(* IEC 61131-3 sources: llm-plc-st-eval/data/processed_definitivo/gemini-3.1-pro-preview/I8/zero_shot, 3 files *)

(* ---- ejec_1.st ---- *)
FUNCTION_BLOCK FB_Compresor
VAR_INPUT
    pOilOk    : BOOL; // Presión de aceite correcta
    tempOk    : BOOL; // Temperatura correcta
    sinAlm    : BOOL; // Ausencia de alarmas
    btnMarcha : BOOL; // Botón de arranque
    btnParo   : BOOL; // Botón de detención
END_VAR

VAR_OUTPUT
    comp         : BOOL; // Comando de marcha del compresor
    causaBloqueo : INT;  // Código del permisivo faltante (0=Ninguno, 1=Aceite, 2=Temp, 3=Alarma)
END_VAR

VAR
    timerOil   : TON;    // Temporizador para validar la presión de aceite
    edgeMarcha : R_TRIG; // Detector de flanco de subida para el botón de marcha
    permisivos : BOOL;   // Bandera interna de todos los permisivos OK
END_VAR

// 1. Evaluación del tiempo de la presión de aceite (3 segundos continuos)
timerOil(IN := pOilOk, PT := T#3S);

// 2. Determinación de la causa de bloqueo (Prioridad al número menor)
IF NOT timerOil.Q THEN
    causaBloqueo := 1; // Falta presión de aceite o no ha transcurrido el tiempo
ELSIF NOT tempOk THEN
    causaBloqueo := 2; // Falta temperatura correcta
ELSIF NOT sinAlm THEN
    causaBloqueo := 3; // Presencia de alarma
ELSE
    causaBloqueo := 0; // Todos los permisivos se cumplen
END_IF;

// 3. Consolidación de permisivos
permisivos := (causaBloqueo = 0);

// 4. Detección de la pulsación de marcha (transición FALSE a TRUE)
edgeMarcha(CLK := btnMarcha);

// 5. Lógica de arranque y paro del compresor
// El paro y la pérdida de permisivos tienen prioridad absoluta
IF btnParo OR NOT permisivos THEN
    comp := FALSE;
// Solo arranca con un nuevo flanco de subida si los permisivos están listos
ELSIF edgeMarcha.Q AND permisivos THEN
    comp := TRUE;
END_IF;

END_FUNCTION_BLOCK

(* ---- ejec_2.st ---- *)
FUNCTION_BLOCK FB_Compresor
VAR_INPUT
    pOilOk    : BOOL; // Presión de aceite correcta
    tempOk    : BOOL; // Temperatura correcta
    sinAlm    : BOOL; // Ausencia de alarmas
    btnMarcha : BOOL; // Botón de arranque
    btnParo   : BOOL; // Botón de parada
END_VAR

VAR_OUTPUT
    comp         : BOOL; // Comando de arranque del compresor
    causaBloqueo : INT;  // Código del permisivo faltante (0=Ninguno, 1=Aceite, 2=Temp, 3=Alarma)
END_VAR

VAR
    tonOil     : TON;    // Temporizador para validar la presión de aceite
    trigMarcha : R_TRIG; // Detector de flanco de subida para el arranque
    permisivos : BOOL;   // Marca interna de todos los permisivos cumplidos
END_VAR

// 1. Temporizador: requiere 3 segundos continuos de pOilOk
tonOil(IN := pOilOk, PT := T#3S);

// 2. Lógica de diagnóstico de bloqueo (prioridad al número menor mediante IF-ELSIF)
IF NOT tonOil.Q THEN
    causaBloqueo := 1; // Falla 1: Presión de aceite no establecida
ELSIF NOT tempOk THEN
    causaBloqueo := 2; // Falla 2: Temperatura incorrecta
ELSIF NOT sinAlm THEN
    causaBloqueo := 3; // Falla 3: Alarma activa
ELSE
    causaBloqueo := 0; // Sin fallas: Todos los permisivos OK
END_IF;

// 3. Evaluación global de permisivos
permisivos := (causaBloqueo = 0);

// 4. Detección de pulsación (transición FALSE a TRUE) del botón de marcha
trigMarcha(CLK := btnMarcha);

// 5. Lógica de control de marcha/paro del compresor
IF btnParo OR NOT permisivos THEN
    // El paro y la pérdida de permisivos tienen prioridad y detienen el equipo
    comp := FALSE;
ELSIF trigMarcha.Q AND permisivos THEN
    // Solo arranca con un nuevo flanco de subida si los permisivos están listos
    comp := TRUE;
END_IF;

END_FUNCTION_BLOCK

(* ---- ejec_3.st ---- *)
FUNCTION_BLOCK FB_Compresor
VAR_INPUT
    pOilOk    : BOOL; // Presión de aceite correcta
    tempOk    : BOOL; // Temperatura correcta
    sinAlm    : BOOL; // Ausencia de alarmas
    btnMarcha : BOOL; // Botón de arranque
    btnParo   : BOOL; // Botón de detención
END_VAR

VAR_OUTPUT
    comp         : BOOL; // Comando de marcha del compresor
    causaBloqueo : INT;  // Indicador del permisivo faltante (0=OK, 1=Aceite, 2=Temp, 3=Alarma)
END_VAR

VAR
    tonOil      : TON;    // Temporizador para validar la presión de aceite
    rTrigMarcha : R_TRIG; // Detector de flanco de subida para el botón de marcha
    permisivos  : BOOL;   // Estado de todos los permisivos combinados
END_VAR

// 1. Evaluación del permisivo de aceite (3 segundos continuos)
tonOil(IN := pOilOk, PT := T#3S);

// 2. Detección de la pulsación de marcha (transición FALSE -> TRUE)
rTrigMarcha(CLK := btnMarcha);

// 3. Lógica de diagnóstico de bloqueo (prioridad al número menor)
IF NOT tonOil.Q THEN
    causaBloqueo := 1; // Falta presión de aceite (o no ha cumplido el tiempo)
ELSIF NOT tempOk THEN
    causaBloqueo := 2; // Falta temperatura correcta
ELSIF NOT sinAlm THEN
    causaBloqueo := 3; // Alarma activa
ELSE
    causaBloqueo := 0; // Todos los permisivos se cumplen
END_IF;

// 4. Agrupación de permisivos
permisivos := (causaBloqueo = 0);

// 5. Lógica de control de marcha/paro del compresor
// El paro y la pérdida de permisivos tienen prioridad absoluta
IF btnParo OR NOT permisivos THEN
    comp := FALSE;
// Solo arranca con el flanco de subida si los permisivos están listos
ELSIF rTrigMarcha.Q AND permisivos THEN
    comp := TRUE;
END_IF;

END_FUNCTION_BLOCK
